// TIA Portal V21 export
// export: Created 2026-08-21T20:18:51.9763251Z, ExportSetting None, DisplayName Totally Integrated Automation Portal, DisplayVersion V21, DisplayName STEP 7 Professional, DisplayVersion V21, DisplayName STEP 7 Safety, DisplayVersion V21, DisplayName Tech WebApplication, DisplayVersion V21, DisplayName WinCC Basic/Comfort/Advanced, DisplayVersion V21, DisplayName WinCC Professional, DisplayVersion V21, DisplayName WinCC Unified, DisplayVersion V21
DATA_BLOCK "ProcessValues_DB"   // DB34
AUTHOR : Siemens AG
FAMILY : ServiceControl
VERSION : 1.0
// stored: InstanceOfName ProcessValues, InstanceOfType FB
"ProcessValues"
   // VAR_INPUT
   //    ProcessValueOutAnalogIn { ExternalAccessible := 'False'; ExternalVisible := 'False'; ExternalWritable := 'False'} : Array[0..0] of "UDT_MTP_AnaProcessValueOut";
   //    ProcessValueOutDigitalIn { ExternalAccessible := 'False'; ExternalVisible := 'False'; ExternalWritable := 'False'} : Array[0..0] of "UDT_MTP_DIntProcessValueOut";
   //    ProcessValueOutBinaryIn { ExternalAccessible := 'False'; ExternalVisible := 'False'; ExternalWritable := 'False'} : Array[0..0] of "UDT_MTP_BinProcessValueOut";
   //    ProcessValueOutStringIn { ExternalAccessible := 'False'; ExternalVisible := 'False'; ExternalWritable := 'False'} : Array[0..0] of "UDT_MTP_StringProcessValueOut";
   //    ProcessValueInAnalogApply { ExternalAccessible := 'False'; ExternalVisible := 'False'; ExternalWritable := 'False'} : Array[0..0] of "UDT_Service_ProcessValueInApply";
   //    ProcessValueInDigitalApply { ExternalAccessible := 'False'; ExternalVisible := 'False'; ExternalWritable := 'False'} : Array[0..0] of "UDT_Service_ProcessValueInApply";
   // END_VAR
   // VAR_OUTPUT
   //    ProcessValueInAnalogOut { ExternalAccessible := 'False'; ExternalVisible := 'False'; ExternalWritable := 'False'} : Array[0..0] of "UDT_MTP_AnaProcessValueOut";
   //    ProcessValueInDigitalOut { ExternalAccessible := 'False'; ExternalVisible := 'False'; ExternalWritable := 'False'} : Array[0..0] of "UDT_MTP_DIntProcessValueOut";
   //    ProcessValueInBinaryOut { ExternalAccessible := 'False'; ExternalVisible := 'False'; ExternalWritable := 'False'} : Array[0..0] of "UDT_MTP_BinProcessValueOut";
   //    ProcessValueInStringOut { ExternalAccessible := 'False'; ExternalVisible := 'False'; ExternalWritable := 'False'} : Array[0..0] of "UDT_MTP_StringProcessValueOut";
   // END_VAR
   // VAR
   //    MTPAnalogIn : Array[0..1] of "UDT_MTP_AnaProcessValueIn";
   //    MTPDigitalIn : Array[0..0] of "UDT_MTP_DIntProcessValueIn";
   //    MTPBinaryIn : Array[0..1] of "UDT_MTP_BinProcessValueIn";
   //    MTPStringIn : Array[0..0] of "UDT_MTP_StringProcessValueIn";
   //    AnalogIn { ExternalAccessible := 'False'; ExternalVisible := 'False'; ExternalWritable := 'False'; S7_SetPoint := 'True'} : Array[0..0] of "ProcessValueInAnalog";
   //    DigitalIn { ExternalAccessible := 'False'; ExternalVisible := 'False'; ExternalWritable := 'False'; S7_SetPoint := 'True'} : Array[0..0] of "ProcessValueInDigital";
   //    BinaryIn { ExternalAccessible := 'False'; ExternalVisible := 'False'; ExternalWritable := 'False'; S7_SetPoint := 'True'} : Array[0..0] of "ProcessValueInBinary";
   //    StringIn { ExternalAccessible := 'False'; ExternalVisible := 'False'; ExternalWritable := 'False'; S7_SetPoint := 'True'} : Array[0..0] of "ProcessValueInString";
   //    MTPAnalogOut : Array[0..1] of "UDT_MTP_AnaProcessValueOut";
   //    MTPDigitalOut : Array[0..0] of "UDT_MTP_DIntProcessValueOut";
   //    MTPBinaryOut : Array[0..0] of "UDT_MTP_BinProcessValueOut";
   //    MTPStringOut : Array[0..0] of "UDT_MTP_StringProcessValueOut";
   //    AnalogOut { ExternalAccessible := 'False'; ExternalVisible := 'False'; ExternalWritable := 'False'; S7_SetPoint := 'True'} : Array[0..0] of "ProcessValueOutAnalog";
   //    DigitalOut { ExternalAccessible := 'False'; ExternalVisible := 'False'; ExternalWritable := 'False'; S7_SetPoint := 'True'} : Array[0..0] of "ProcessValueOutDigital";
   //    BinaryOut { ExternalAccessible := 'False'; ExternalVisible := 'False'; ExternalWritable := 'False'; S7_SetPoint := 'True'} : Array[0..0] of "ProcessValueOutBinary";
   //    StringOut { ExternalAccessible := 'False'; ExternalVisible := 'False'; ExternalWritable := 'False'; S7_SetPoint := 'True'} : Array[0..0] of "ProcessValueOutString";
   // END_VAR
BEGIN
   MTPAnalogIn[0].V := 1500.0;
   MTPAnalogIn[0].SclMinCur := 0.0;
   MTPAnalogIn[0].SclMaxCur := 3000.0;
   MTPAnalogIn[0].UnitCur := 1038;
   MTPAnalogIn[0].SclMinExt := 0.0;
   MTPAnalogIn[0].SclMaxExt := 3000.0;
   MTPAnalogIn[0].UnitExt := 1038;
   MTPBinaryIn[0].V := True;
   MTPBinaryIn[0].VState0 := 'Valve next PEA c';
   MTPBinaryIn[0].VState1 := 'Valve next PEA o';
   MTPAnalogOut[0..1].V := 0.0;
   MTPAnalogOut[0..1].VSclMin := 0.0;
   MTPAnalogOut[0..1].VSclMax := 32.0;
   MTPAnalogOut[0].VUnit := 1351;
   MTPAnalogOut[1].VUnit := 1322;
END_DATA_BLOCK
